FUNCTION_BLOCK FB_Palletizer IMPLEMENTS ITF_Palletizer
VAR_INPUT
END_VAR
VAR_OUTPUT
END_VAR
VAR
END_VAR

{warning 'Add method implementation '}
METHOD Aborted : BOOL
END_METHOD

{warning 'Add method implementation '}
METHOD Aborting : BOOL
END_METHOD

{warning 'Add method implementation '}
METHOD Clearing : BOOL
END_METHOD

{warning 'Add method implementation '}
METHOD Execute : BOOL
END_METHOD

{warning 'Add method implementation '}
METHOD Held : BOOL
END_METHOD

{warning 'Add method implementation '}
METHOD Holding : BOOL
END_METHOD

{warning 'Add method implementation '}
METHOD Idle : BOOL
END_METHOD

{warning 'Add method implementation '}
METHOD Resetting : BOOL
END_METHOD

{warning 'Add method implementation '}
METHOD Starting : BOOL
END_METHOD

{warning 'Add method implementation '}
METHOD Stopped : BOOL
END_METHOD

{warning 'Add method implementation '}
METHOD Stopping : BOOL
END_METHOD

{warning 'Add method implementation '}
METHOD Suspended : BOOL
END_METHOD

{warning 'Add method implementation '}
METHOD Suspending : BOOL
END_METHOD

{warning 'Add method implementation '}
METHOD Unholding : BOOL
END_METHOD

{warning 'Add method implementation '}
METHOD Unsuspending : BOOL
END_METHOD

END_FUNCTION_BLOCK

(* stored: Version 1.1.0.1
   POU FB_Palletizer: Id {6bcdea34-befa-4851-b701-54154571fa23}, SpecialFunc None
   Folder Methods: Id {328a659f-6935-4661-bc18-54b0fa869ace}
   Method Aborted: Id {3eb12933-a46e-4508-b1b1-d7c960fc3d26}
   Method Aborting: Id {d12fdfca-5fe1-4054-b56d-d9e0ff65597e}
   Method Clearing: Id {90e5dfd0-9549-4982-b0a1-ac32ba1e6292}
   Method Execute: Id {28a22277-8a7e-4bd6-bec1-78218065b663}
   Method Held: Id {fc6bf354-b8db-41cb-a7ec-f7251ff0298e}
   Method Holding: Id {a7aec294-162a-4b83-9988-b8f31c4751a2}
   Method Idle: Id {39494d41-c348-475d-b27a-e70f1e0665a8}
   Method Resetting: Id {fe910404-29f4-40cc-b9da-ffcee1e49c0c}
   Method Starting: Id {d2a787b4-56af-4df8-93c0-3884d94a0e09}
   Method Stopped: Id {c7a431f7-6769-4be9-aa5f-f8acf4378890}
   Method Stopping: Id {59a02c41-e1b1-466e-9b53-10d0802d9340}
   Method Suspended: Id {fe3f7e2b-bbd4-41e2-bfeb-7bcdbec906bf}
   Method Suspending: Id {e179ce52-3b13-4be4-9f35-965df06c3c24}
   Method Unholding: Id {7e41c785-9fe6-4c55-8866-22120e934b35}
   Method Unsuspending: Id {c447ee90-96bc-4841-aa23-a54cffbc916b} *)
